// TIA Portal V20 export
// export: Created 2026-10-20T18:56:03.5836865Z, ExportSetting None, DisplayName Totally Integrated Automation Portal, DisplayVersion V20 Update 6, DisplayName TIA Portal Openness, DisplayVersion V20 Update 6, DisplayName TIA Portal Version Control Interface, DisplayVersion V20 Update 6, DisplayName SINAMICS Startdrive Advanced, DisplayVersion V20 SP1, DisplayName SINAMICS Startdrive G130, G150, S120, S150, SINAMICS MV, G220, S200, S210, DisplayVersion V20 SP1, DisplayName SINAMICS Startdrive G110M, G120, G120C, G120D, G120P, G115D, DisplayVersion V20 SP1, DisplayName STEP 7 Professional, DisplayVersion V20 Update 6, DisplayName STEP 7 Safety, DisplayVersion V20 Update 2, DisplayName WinCC Basic/Comfort/Advanced, DisplayVersion V20 Update 6, DisplayName WinCC Unified, DisplayVersion V20 Update 6
VAR_GLOBAL   // PLC tag table "Lock_12"
   "Lock Reset_12" AT %Q1508.0 : Bool;
   Lamps_12 AT %QB1506 : Byte;
   Switches_12 AT %IB1855 : Byte;
   Lock_12_Closed_CH2 AT %I1847.1 : Bool;
   "Solenoid Enable_12" AT %Q1507.0 : Bool;
   Lock_12_Estop_CH2 AT %I1847.3 : Bool;
   Lock_12_Closed_CH1 AT %I1847.0 : Bool;
   Lock_12_Estop_CH1 AT %I1847.2 : Bool;
   Lock_12_Reset_Input4 AT %Q1848.3 : Bool;
   Lock_12_Reset_Input2 AT %Q1848.1 : Bool;
   Lock_12_Reset_Input1 AT %Q1848.0 : Bool;
   Lock_12_Reset_Input3 AT %Q1848.2 : Bool;
   "Guard Position_12" AT %I1856.0 : Bool;
   "Lock Position_12" AT %I1857.0 : Bool;
END_VAR
